Fanuc KAREL source: kt00475.KL

-- PROVISIONAL review KL for V770-1; original PC SHA256 0b6df09d993100a74f02f448ea1b5e694e33dc5569074a4fe4d76a74e35a0833
-- Incomplete behavior may be omitted. Consult companion uncertainty JSON. Do not deploy.
PROGRAM KT00475
%NOLOCKGROUP
-- UNRESOLVED_DECL P1 type=000101
-- UNRESOLVED_DECL P2 type=000101
-- UNRESOLVED_DECL OUT type=000102
BEGIN
  -- UNRESOLVED_PC offsets 5-34; opcodes 49,49,60,7E,4A
  -- UNRESOLVED_PC offsets 39-43; opcodes 7F
END KT00475
